TYPE "ST_ModelId"
VERSION : 0.1
   STRUCT
      "ModelCode" : String[64];
      "Family" : String[64];
      "Variant" : String[64];
      "Fields" : Array[1..8] of "ST_ModelField";
      "NField" : Int;
   END_STRUCT;
END_TYPE
